// TIA Portal V20 export
Screen "StyleWrite"  1276x673
  ScreenItem "线_1" at 0,85 size 1360x2  Type=HmiLine
  ScreenItem "符号 IO 域_1" at 454,39 size 500x42  Type=HmiSymbolicIOField
  ScreenItem "Button_Special_2" at 1086,8 size 90x60  Type=HmiButton
  ScreenItem "Button_Special_3" at 1178,8 size 90x60  Type=HmiButton
  ScreenItem "permanentareaborderrectangle" at 0,0 size 0x0  Type=HmiRectangle
  ScreenItem "Button_Back" at 6,8 size 90x60  Type=HmiButton
  ScreenItem "Title_OPMode1_ScreenOverview_X390_Y2" at 454,7 size 500x30  Type=HmiTextBox
  ScreenItem "Faceplate container_1" at 74,87 size 1119x584  Type=HmiFaceplateContainer
